Fanuc KAREL source: KS00004.KL

PROGRAM KS00004
%NOLOCKGROUP
TYPE
  REC_T = STRUCTURE
    VALUE: INTEGER
    FLAG: BOOLEAN
  ENDSTRUCTURE
VAR
  A: REC_T
  B: REC_T
  FLAG: BOOLEAN
  N: INTEGER
  STATUS: INTEGER
  PN: STRING[80]
  VN: STRING[80]
BEGIN
  PN = ''
  VN = 'A'
  FLAG = UNINIT(A)
END KS00004
